// TIA Portal V21 export
ScreenTemplate "Tpl"  NonexNone
  ScreenLayer 
